TYPE ST_SpindlePDSXLA170ClutchStatus_1 :
STRUCT
	bRotatingS1					:BOOL;						(* Spindle rotating S1 *)
	bToolNotClampedS2			:BOOL;						(* Tool not clamped S2 *)
	bToolPresentS3				:BOOL;						(* Tool present S3 *)
	bClutchInBaseS4				:BOOL;						(* Clutch in base position S4 *)
END_STRUCT
END_TYPE

(* stored: Version 1.1.0.1, ProductVersion 3.1.4024.15
   DUT ST_SpindlePDSXLA170ClutchStatus_1: Id {0292834f-aca6-4416-a9a3-96d1ffaedd79} *)
